// Generated by voz_llm_plc_agent
// Target: Siemens TIA Portal V18 - SCL external source
// Review and compile before any download to physical hardware.

FUNCTION_BLOCK "PLC_PRG"
{ S7_Optimized_Access := 'TRUE' }
VERSION : 0.1
VAR_INPUT
   I_Piece_Sensor : Bool := FALSE;
   I_Emergency : Bool := FALSE;
   I_Start : Bool := FALSE;
END_VAR
VAR_OUTPUT
   Q_Alarm : Bool := FALSE;
END_VAR
VAR
   T_SensorTimeout {InstructionName := 'TON_TIME'; LibVersion := '1.0'} : TON_TIME;
   M_SensorLastState : Bool;
   M_SupervisionActive : Bool;
END_VAR
BEGIN
(* Supervision del sensor desde la orden de arranque: alarma si no cambia de estado durante el *)
(* tiempo indicado; cada cambio reinicia la cuenta. *)
IF FALSE OR #I_Emergency THEN
    #M_SupervisionActive := FALSE;
ELSIF #I_Start THEN
    #M_SupervisionActive := TRUE;
END_IF;

#T_SensorTimeout(IN := #M_SupervisionActive AND (#I_Piece_Sensor = #M_SensorLastState) AND NOT #I_Emergency, PT := T#5s);
#Q_Alarm := #T_SensorTimeout.Q AND #M_SupervisionActive AND NOT #I_Emergency;
#M_SensorLastState := #I_Piece_Sensor;
END_FUNCTION_BLOCK

DATA_BLOCK "DB_PLC_PRG"
{ S7_Optimized_Access := 'TRUE' }
VERSION : 0.1
NON_RETAIN
"PLC_PRG"
BEGIN
END_DATA_BLOCK

ORGANIZATION_BLOCK "Main"
{ S7_Optimized_Access := 'TRUE' }
VERSION : 0.1
BEGIN
   "DB_PLC_PRG"(
      I_Piece_Sensor := "I_Piece_Sensor",
      I_Emergency := "I_Emergency",
      Q_Alarm => "Q_Alarm",
      I_Start := "I_Start"
   );
END_ORGANIZATION_BLOCK
